Fanuc KAREL source: kt00489.KL

PROGRAM KT00489
%STACKSIZE=65535
%PRIORITY=65535
%NOLOCKGROUP
VAR
P1 : POSITION
P2 : JOINTPOS9
OUT : POSITION
BEGIN
-- UNRESOLVED_PC line 8 opcodes [49 49 7E 60 4A] marker_code=0
END KT00489
